// TIA Portal V21 export
TYPE "AxisAS_CFG_Type_v4"
// Configurazione asse AxisAS_Mng_v4
   STRUCT
      fMaxSpeed { S7_SetPoint := 'True'} : Real := 100.0;   // Limite SUP velocità richiesta (mm/s)
      fMinSpeed { S7_SetPoint := 'True'} : Real := 5.0;   // Velocità minima di accostamento e correzione finale (mm/s), deve essere > 0
      fMinAccRamp { S7_SetPoint := 'True'} : Real := 100.0;   // Limite INF accelerazione (mm/s^2)
      fMaxAccRamp { S7_SetPoint := 'True'} : Real := 1200.0;   // Limite SUP accelerazione (mm/s^2)
      fMinDecRamp { S7_SetPoint := 'True'} : Real := 100.0;   // Limite INF decelerazione (mm/s^2)
      fMaxDecRamp { S7_SetPoint := 'True'} : Real := 800.0;   // Limite SUP decelerazione (mm/s^2)
      fJerk { S7_SetPoint := 'True'} : Real := 0.0;   // Jerk (mm/s^3): 0 = trapezio puro. Valori tipici 5..10 x accelerazione per un profilo morbido
      fThreshold_SUP_AutoSpeed { S7_SetPoint := 'True'} : Real := 500.0;   // Autospeed: distanza oltre la quale si usa la velocità richiesta (mm)
      fThreshold_INF_AutoSpeed { S7_SetPoint := 'True'} : Real := 0.0;   // Autospeed: distanza a cui corrisponde fMinSpeed (mm)
      fMotWindPos { S7_SetPoint := 'True'} : Real := 1.0;   // Finestra di posizione per In posizione (mm), deve essere > 0
      fMotWindPosBig { S7_SetPoint := 'True'} : Real := 30.0;   // Finestra allargata di posizione (mm)
      fMotWindSpeed { S7_SetPoint := 'True'} : Real := 10.0;   // Velocità reale massima per considerare il motore fermo (mm/s)
      fMotAdvStopPosition { S7_SetPoint := 'True'} : Real := 0.0;   // Anticipo (+) / ritardo (-) inizio decelerazione (mm): compensa inerzie e ritardi
      tAdvStop { S7_SetPoint := 'True'} : Time := T#0ms;   // Compensazione inerzia: ritardo tra riferimento e velocità reale. Anticipa decelerazione e arresto in proporzione alla velocità
      fReposWindow { S7_SetPoint := 'True'} : Real := 0.0;   // Riposizionamento automatico da fermo se l'encoder esce da questa finestra (mm). 0=disabilitato
      xPosLoop { S7_SetPoint := 'True'} : Bool := false;   // =1 il motore insegue l'asse virtuale (tempi ripetibili, coordinamento assi). =0 solo profilo, decisioni su encoder
      fKp_Pos { S7_SetPoint := 'True'} : Real := 2.0;   // xPosLoop: guadagno proporzionale sull'errore di inseguimento (1/s)
      fKp_PosDec { S7_SetPoint := 'True'} : Real := 0.0;   // xPosLoop: guadagno aggiunto a piramide (1/s), cresce da 0 a fKp_PosDec mentre la velocità scende dal massimo del movimento (come fKPpidDec_Pos v2.0). 0 = disabilitato
      fPosLoopLimitPct { S7_SetPoint := 'True'} : Real := 20.0;   // xPosLoop: limite della correzione in % di fMaxSpeed
      fMaxErrEnc { S7_SetPoint := 'True'} : Real := 20.0;   // xPosLoop: errore di inseguimento massimo per allarme (mm). 0 = allarme disabilitato
      fJogSpeed { S7_SetPoint := 'True'} : Real := 10.0;   // Velocità JOG (mm/s)
      fJogAcc { S7_SetPoint := 'True'} : Real := 10.0;   // Accelerazione JOG (mm/s^2)
      fJogDec { S7_SetPoint := 'True'} : Real := 10.0;   // Decelerazione JOG (mm/s^2)
      fOffSResLevel { S7_SetPoint := 'True'} : Real := 50.0;   // Ricerca livello: anticipo per raggiungere la velocità di ricerca prima della quota di inizio (50 se mm, 5 se gradi)
      tBrakeDelay_Fwd { S7_SetPoint := 'True'} : Time := T#100ms;   // Ritardo chiusura freno a fine movimento avanti/salita
      tBrakeDelay_Bkw { S7_SetPoint := 'True'} : Time := T#100ms;   // Ritardo chiusura freno a fine movimento indietro/discesa
      tDriveOnReq { S7_SetPoint := 'True'} : Time := T#5s;   // Mantenimento marcia (inverter magnetizzato) dopo l'arresto
      tDriveReadyTimeout { S7_SetPoint := 'True'} : Time := T#3s;   // Tempo massimo di attesa inverter pronto/magnetizzato
      tCtrEndPos { S7_SetPoint := 'True'} : Time := T#3s;   // Tempo massimo per entrare in posizione dall'arrivo in finestra. T#0s = disabilitato
      tStallTime { S7_SetPoint := 'True'} : Time := T#2s;   // Allarme asse bloccato: motore comandato ma encoder fermo o in senso opposto. T#0s = disabilitato
   END_STRUCT;
END_TYPE
